(* IEC 61131-3 sources: Gen-AI/release/member2-v1.1/成员2_提交包_v1.1/validation/toolchain_smoke_v1.1/C00_good/tools/check/authoritative, 1 file *)

(* ---- source.st ---- *)
FUNCTION_BLOCK FB_AgentProbeGood
VAR_INPUT
 x : BOOL;
END_VAR
VAR_OUTPUT
 y : BOOL;
END_VAR
y := x;
END_FUNCTION_BLOCK
